TYPE ST_Parameter :
STRUCT
	fPosition: LREAL;
	fVelocity: LREAL;
	fAcceleration: LREAL;
	fDeceleration: LREAL;
	fJerk: LREAL;
END_STRUCT
END_TYPE

(* stored: Version 1.1.0.1, ProductVersion 3.1.4024.12
   DUT ST_Parameter: Id {9997025b-dcf0-4adf-80d7-0ea551e3deed} *)
